// TIA Portal V21 export
// export: Created 2026-10-14T03:06:09.1558359Z, ExportSetting WithDefaults, DisplayName Totally Integrated Automation Portal, DisplayVersion V21, DisplayName STEP 7 Professional, DisplayVersion V21, DisplayName STEP 7 Safety, DisplayVersion V21, DisplayName Tech WebApplication, DisplayVersion V21, DisplayName WinCC Basic/Comfort/Advanced, DisplayVersion V21, DisplayName WinCC Unified, DisplayVersion V21
VAR_GLOBAL   // PLC tag table "DemocaseAppTagTable"
   ControlUnit_AddressIn AT %I300.0 : "PD_TEL_393_IN";
   ControlUnit_AddressOut AT %Q300.0 : "PD_TEL_393_OUT";
   ET200_AI_0 AT %IW2 : Int;
   ET200_AI_1 AT %IW4 : Int;
   OutputCam_1_Interface_Address AT %Q303.5 : Bool;
   TB30_AI_0 AT %IW342 : Word;
   TB30_AI_1 AT %IW344 : Word;
END_VAR
